// TIA Portal V19 export
// export: Created 2026-10-15T10:10:17.3827368Z, ExportSetting WithDefaults, DisplayName Totally Integrated Automation Portal, DisplayVersion V19, DisplayName TIA Portal Openness, DisplayVersion V19, DisplayName TIA Portal Version Control Interface, DisplayVersion V19, DisplayName STEP 7 Professional, DisplayVersion V19, DisplayName STEP 7 Safety, DisplayVersion V19, DisplayName WinCC Basic/Comfort/Advanced, DisplayVersion V19, DisplayName WinCC Unified, DisplayVersion V19
DATA_BLOCK "ROLL_DB19"   // DB5
{ S7_Optimized_Access := 'TRUE' }
VERSION : 0.1
// stored: AutoNumber true, DBAccessibleFromOPCUA true, DBAccessibleFromWebserver true, IsOnlyStoredInLoadMemory false, IsRetainMemResEnabled false, IsWriteProtectedInAS false, MemoryReserve 100
   VAR RETAIN
      DW : Array[0..131] of Word;
   END_VAR
BEGIN
   DW[0] := WORD#16#FFFF;
   DW[1] := WORD#16#0020;
   DW[2] := WORD#16#0014;
   DW[3..127] := WORD#16#FFFF;
   DW[128..129] := WORD#16#0001;
   DW[130] := WORD#16#0020;
END_DATA_BLOCK
